(* IEC 61131-3 sources: llm-plc-st-eval/data/processed_definitivo/qwen2.5-coder_14b/C4/few_shot, 3 files *)

(* ---- ejec_1.st ---- *)
FUNCTION_BLOCK FB_D
VAR_INPUT
    demanda : BOOL; (* Indica si hay una demanda de activación *)
    falla1 : BOOL;  (* Indica si hay una falla en el sistema 1 *)
    falla2 : BOOL;  (* Indica si hay una falla en el sistema 2 *)
END_VAR
VAR_OUTPUT
    bomba1 : BOOL;  (* Controla la activación de la bomba 1 *)
    bomba2 : BOOL;  (* Controla la activación de la bomba 2 *)
    almFalla : BOOL; (* Almacena el estado de la última falla detectada *)
END_VAR
VAR
    turno : BOOL;   (* Variable de estado para alternar entre bombas *)
    fDem : R_TRIG;  (* Detector de flanco de subida en la demanda *)
END_VAR

(* Detecta el flanco de subida en la demanda *)
fDem(CLK := demanda);

(* Cambia el turno entre bombas cuando hay una demanda *)
IF fDem.Q THEN
    turno := NOT turno;
END_IF

(* Control de las bombas y almacenamiento de la última falla *)
IF demanda THEN
    IF turno THEN
        bomba1 := NOT falla1; (* Activa bomba1 si no hay falla1 *)
        bomba2 := falla1 AND NOT falla2; (* Activa bomba2 si hay falla1 y no hay falla2 *)
        almFalla := falla1; (* Almacena el estado de falla1 *)
    ELSE
        bomba2 := NOT falla2; (* Activa bomba2 si no hay falla2 *)
        bomba1 := falla2 AND NOT falla1; (* Activa bomba1 si hay falla2 y no hay falla1 *)
        almFalla := falla2; (* Almacena el estado de falla2 *)
    END_IF
ELSE
    bomba1 := FALSE; (* Desactiva bomba1 si no hay demanda *)
    bomba2 := FALSE; (* Desactiva bomba2 si no hay demanda *)
    almFalla := FALSE; (* Limpia el registro de falla *)
END_IF
END_FUNCTION_BLOCK

(* ---- ejec_2.st ---- *)
FUNCTION_BLOCK FB_D
VAR_INPUT
    demanda : BOOL; (* Indica si hay una demanda de activación *)
    falla1 : BOOL; (* Indica si la bomba1 está fallando *)
    falla2 : BOOL; (* Indica si la bomba2 está fallando *)
END_VAR
VAR_OUTPUT
    bomba1 : BOOL; (* Control de la bomba1 *)
    bomba2 : BOOL; (* Control de la bomba2 *)
    almFalla : BOOL; (* Almacena la última falla detectada *)
END_VAR
VAR
    turno : BOOL; (* Variable de control para alternar entre bomba1 y bomba2 *)
    fDem : R_TRIG; (* Flanco de subida de la demanda *)
END_VAR

(* Detecta el flanco de subida de la demanda *)
fDem(CLK := demanda);
IF fDem.Q THEN
    (* Alterna el turno entre bomba1 y bomba2 *)
    turno := NOT turno;
END_IF

(* Si hay una demanda *)
IF demanda THEN
    (* Si el turno está en bomba1 *)
    IF turno THEN
        (* Activa bomba1 si no está fallando *)
        bomba1 := NOT falla1;
        (* Activa bomba2 si está fallando bomba1 y no está fallando bomba2 *)
        bomba2 := falla1 AND NOT falla2;
        (* Almacena la última falla detectada *)
        almFalla := falla1;
    ELSE
        (* Si el turno está en bomba2 *)
        (* Activa bomba2 si no está fallando *)
        bomba2 := NOT falla2;
        (* Activa bomba1 si está fallando bomba2 y no está fallando bomba1 *)
        bomba1 := falla2 AND NOT falla1;
        (* Almacena la última falla detectada *)
        almFalla := falla2;
    END_IF
ELSE
    (* Si no hay demanda, apaga ambas bombas *)
    bomba1 := FALSE;
    bomba2 := FALSE;
    (* Limpia el registro de la última falla *)
    almFalla := FALSE;
END_IF
END_FUNCTION_BLOCK

(* ---- ejec_3.st ---- *)
FUNCTION_BLOCK FB_D
VAR_INPUT
    demanda : BOOL; (* Señal de demanda para activar una bomba *)
    falla1 : BOOL; (* Indica una falla en la bomba 1 *)
    falla2 : BOOL; (* Indica una falla en la bomba 2 *)
END_VAR
VAR_OUTPUT
    bomba1 : BOOL; (* Control de la bomba 1 *)
    bomba2 : BOOL; (* Control de la bomba 2 *)
    almFalla : BOOL; (* Almacena la información de la última falla detectada *)
END_VAR
VAR
    turno : BOOL; (* Variable de estado para alternar entre bomba1 y bomba2 *)
    fDem : R_TRIG; (* Temporizador de flanco ascendente para detectar demanda *)
END_VAR

(* Configura el temporizador de flanco ascendente con la señal de demanda *)
fDem(CLK := demanda);

(* Si se detecta una demanda (flanco ascendente) *)
IF fDem.Q THEN
    (* Alterna el estado de la variable turno *)
    turno := NOT turno;
END_IF

(* Si hay una demanda *)
IF demanda THEN
    (* Si el turno está en TRUE *)
    IF turno THEN
        (* Activa bomba1 si no hay falla en bomba1 *)
        bomba1 := NOT falla1;
        (* Activa bomba2 si hay falla en bomba1 y no hay falla en bomba2 *)
        bomba2 := falla1 AND NOT falla2;
        (* Almacena la información de la última falla detectada *)
        almFalla := falla1;
    (* Si el turno está en FALSE *)
    ELSE
        (* Activa bomba2 si no hay falla en bomba2 *)
        bomba2 := NOT falla2;
        (* Activa bomba1 si hay falla en bomba2 y no hay falla en bomba1 *)
        bomba1 := falla2 AND NOT falla1;
        (* Almacena la información de la última falla detectada *)
        almFalla := falla2;
    END_IF
(* Si no hay demanda *)
ELSE
    (* Desactiva ambas bombas *)
    bomba1 := FALSE;
    bomba2 := FALSE;
    (* Limpia la información de la última falla detectada *)
    almFalla := FALSE;
END_IF
END_FUNCTION_BLOCK
